// TIA Portal V21 export
DATA_BLOCK "IDB_Conveyor1200"   // DB1
// stored: InstanceOfName FB_Conveyor1200, InstanceOfType FB
"FB_Conveyor1200"
   // VAR_INPUT
   //    Start : Bool;
   //    Stop : Bool;
   //    SpeedRaw : Int;
   // END_VAR
   // VAR_OUTPUT
   //    Motor : Bool;
   //    Speed : Real;
   //    DelayMilliseconds : DInt;
   // END_VAR
   // VAR
   //    StartDelay { S7_SetPoint := 'True'} : TON_TIME;
   //    Running : Bool;
   // END_VAR
BEGIN
END_DATA_BLOCK
